Fanuc KAREL source: KT00829.KL

PROGRAM KT00829
%NOLOCKGROUP
VAR
  B1: BOOLEAN
  B2: BOOLEAN
  OUT: REAL
BEGIN
  B1 = TRUE
  B2 = FALSE
  B1 = TRUE
  B2 = FALSE
  OUT = SIN(B1)
END KT00829
